(*
SPDX-FileCopyrightText: © 2026 Oleksandr Tiutyk <trofimich@gmail.com>
SPDX-License-Identifier: MIT
License: https://opensource.org/license/mit
*)

(*!
<summary>Orders generic storage lexicographically by bytes and then by size.</summary>
<description>
Non-null addresses must reference readable storage of the declared Size. Two null addresses compare equal; one
null address sorts before a non-null address. Compares the common byte prefix, then Size. TypeClass does not
alter this byte order: string terminators, trailing storage, padding and pointer fields all participate. Use
StringComparer or WStringComparer for terminated-text ordering. OBJECT payload is compared as bytes without
invoking object methods; padding and pointer fields participate. Descriptors are passed by value; payload
remains borrowed and is not modified, cloned, released or retained. IsMemoryOwner does not affect comparison.
</description>
*)

FUNCTION_BLOCK ByteArrayComparer EXTENDS TOF_Core.Object IMPLEMENTS TOF_Core.IComparer
VAR_STAT
	//! <summary>Class name shared by all instances of this function block.</summary>
	{attribute 'hide'}
	_ClassName : STRING := __POUNAME();
END_VAR

{attribute 'monitoring' := 'call'}
PROPERTY ClassName : REFERENCE TO STRING
GET
ClassName REF= _ClassName;
END_GET
END_PROPERTY

(*!
<summary>Compares the first operand with the second using this ordering strategy.</summary>
<description>
Non-null addresses must reference readable storage of the declared Size. Two null addresses compare equal; one
null address sorts before a non-null address. Compares the common byte prefix, then Size. TypeClass does not
alter this byte order: string terminators, trailing storage, padding and pointer fields all participate. Use
StringComparer or WStringComparer for terminated-text ordering. OBJECT payload is compared as bytes without
invoking object methods; padding and pointer fields participate. Descriptors are passed by value; payload
remains borrowed and is not modified, cloned, released or retained. IsMemoryOwner does not affect comparison.
Descendants cannot replace this standard ordering; implement IComparer separately for a different ordering
strategy.
</description>
*)
//!<param name="first">First descriptor; referenced storage is borrowed for the call.</param>
//!<param name="second">Second descriptor; referenced storage is borrowed for the call.</param>
{attribute "object_name" := "Compare"}
METHOD FINAL Compare : TOF_Core.COMPARISON_RESULT
VAR_INPUT
	first : TOF_Core.GENERIC_VALUE;
	second : TOF_Core.GENERIC_VALUE;
END_VAR
VAR
	leftPointer : POINTER TO BYTE;
	rightPointer : POINTER TO BYTE;

	i : ULINT;
	minSize : ULINT;
END_VAR
IF first.Address = 0 AND_THEN second.Address = 0 THEN
	Compare := TOF_Core.COMPARISON_RESULT.FIRST_EQUAL_TO_SECOND;
	RETURN;
END_IF

IF first.Address = 0 THEN
	Compare := TOF_Core.COMPARISON_RESULT.FIRST_LESS_THAN_SECOND;
	RETURN;
END_IF

IF second.Address = 0 THEN
	Compare := TOF_Core.COMPARISON_RESULT.FIRST_GREATER_THAN_SECOND;
	RETURN;
END_IF

minSize := MIN(first.Size, second.Size);

i := 0;

WHILE i < minSize DO
	leftPointer := first.Address + TO_LWORD(i);
	rightPointer := second.Address + TO_LWORD(i);

	IF leftPointer^ < rightPointer^ THEN
		Compare := TOF_Core.COMPARISON_RESULT.FIRST_LESS_THAN_SECOND;
		RETURN;
	ELSIF leftPointer^ > rightPointer^ THEN
		Compare := TOF_Core.COMPARISON_RESULT.FIRST_GREATER_THAN_SECOND;
		RETURN;
	END_IF

	i := i + 1;
END_WHILE

IF first.Size < second.Size THEN
	Compare := TOF_Core.COMPARISON_RESULT.FIRST_LESS_THAN_SECOND;
ELSIF first.Size > second.Size THEN
	Compare := TOF_Core.COMPARISON_RESULT.FIRST_GREATER_THAN_SECOND;
ELSE
	Compare := TOF_Core.COMPARISON_RESULT.FIRST_EQUAL_TO_SECOND;
END_IF
END_METHOD

{attribute 'monitoring' := 'call'}
PROPERTY NamespaceName : REFERENCE TO STRING
GET
NamespaceName REF= CurrentNamespace.Name;
END_GET
END_PROPERTY

{attribute 'monitoring' := 'call'}
PROPERTY SelfSize : ULINT
GET
SelfSize := XSIZEOF(THIS^);
END_GET
END_PROPERTY

END_FUNCTION_BLOCK

(* stored: Version 1.1.0.1
   POU ByteArrayComparer: Id {2bb53bb7-7d07-4a7a-896e-016e853fd868}, SpecialFunc None
   Property ClassName: Id {cf39d53b-ed13-4edf-ad55-696c13de665b}
   Get Get: Id {d30e6779-120e-49c2-abe1-17cbfac7965e}
   Method Compare: Id {ee7448b3-b623-4697-a6c8-19f6c43d07cb}
   Property NamespaceName: Id {9a7e1f84-1d7c-4766-b019-8e9775b5d9ca}
   Get Get: Id {f3eef584-0d20-4a97-ba32-a95b52b6625c}
   Property SelfSize: Id {b1a1240f-8b51-48b9-84a3-3c39c9b5cd85}
   Get Get: Id {7cf65b52-2f9d-4aa5-9cb0-fb0f5d03a50d} *)
